(* IEC 61131-3 sources: ctrlx-ai-coding/skills/ctrlx-opcon-engineering/assets/library-examples/inntai/plc/FB_InntaiWireFixture, 4 files *)

(* ---- Close.st ---- *)
METHOD PUBLIC Close : DINT
(* BODY *)
IF ( NOT _opened )
THEN
  AlreadyClosedCalls := AlreadyClosedCalls + 1;
  Close              := -601;
ELSE
  _opened := FALSE;
  Close   := OK;
END_IF

(* ---- Read.st ---- *)
METHOD PUBLIC Read : DINT
VAR_INPUT
  pData        : POINTER TO BYTE;
  DataLen      : SIZE_T;
  rBytesRead   : REFERENCE TO SIZE_T;
  rReadTimeout : REFERENCE TO BOOL;
END_VAR
VAR
  _chunk : UINT;
  _i     : UINT;
END_VAR
(* BODY *)
_chunk := MIN(TO_UINT(DataLen), MIN(_count, 17));
IF ( _chunk > 0 )
THEN
  FOR _i := 0 TO _chunk - 1
  DO
    pData[_i] := _queue[_i];
  END_FOR
  _count := _count - _chunk;
  IF ( _count > 0 )
  THEN
    FOR _i := 0 TO _count - 1
    DO
      _queue[_i] := _queue[_i + _chunk];
    END_FOR
  END_IF
  ReadChunks   := ReadChunks + 1;
  MaxReadChunk := MAX(MaxReadChunk, _chunk);
END_IF
rBytesRead   := _chunk;
rReadTimeout := ( _chunk = 0 );
Read         := OK;

(* ---- Write.st ---- *)
METHOD PUBLIC Write : DINT
VAR_INPUT
  pData         : POINTER TO BYTE;
  DataLen       : SIZE_T;
  rBytesWritten : REFERENCE TO SIZE_T;
END_VAR
VAR
  _bcc : BYTE;
  _i   : UINT;
END_VAR
(* BODY *)
_bcc := 0;
FOR _i := 0 TO TO_UINT(DataLen) - 2
DO
  _bcc := _bcc XOR pData[_i];
END_FOR
WireValid := WireValid AND ( pData[0] = 2 ) AND
             ( pData[DataLen-2] = 3 ) AND ( _bcc = pData[DataLen-1] );
IF ( NOT WireValid )
THEN
  Write := -10009;
  RETURN;
END_IF
IF ( pData[1] = 82 ) AND
   ( pData[2] = 80 )
THEN
  FOR _i := 0 TO SIZEOF(ReplyParameters) - 1
  DO
    _queue[_i] := ReplyParameters[_i];
  END_FOR
  _count := SIZEOF(ReplyParameters);
ELSIF ( pData[1] = 67 ) AND
      ( pData[2] = 83 )
THEN
  CsCalls := CsCalls + 1;
  FOR _i := 0 TO SIZEOF(ReplyBaseline) - 1
  DO
    IF ( FreshOnRead ) THEN
      _queue[_i] := ReplyFresh[_i];
    ELSE
      _queue[_i] := ReplyBaseline[_i];
    END_IF
  END_FOR
  _count := SIZEOF(ReplyBaseline);
ELSE
  FOR _i := 0 TO SIZEOF(ReplyOk) - 1
  DO
    _queue[_i] := ReplyOk[_i];
  END_FOR
  _count   := SIZEOF(ReplyOk);
  _pending := AutoResult AND ( pData[1] = 83 ) AND ( pData[2] = 84 );
  IF ( pData[1] = 83 ) AND ( pData[2] = 84 ) THEN
    StartCalls := StartCalls + 1;
  END_IF
END_IF
IF ( SuppressReply )
THEN
  _count := 0;
END_IF
rBytesWritten := DataLen;
Write         := OK;

(* ---- Open.st ---- *)
METHOD PUBLIC Open : DINT
VAR_INPUT
  BaudRate  : OC_OpconBaseCommonDef.OpconSerialBaudRate;
  DataFrame : OC_OpconBaseCommonDef.OpconSerialDataFrame;
  Handshake : OC_OpconBaseCommonDef.OpconSerialHandshakeType;
END_VAR
(* BODY *)
ConfigurationCorrect :=
(BaudRate = OC_OpconBaseCommonDef.OpconSerialBaudRate.BAUD_9600) AND
(DataFrame = OC_OpconBaseCommonDef.OpconSerialDataFrame.FRAME_8N1) AND
(Handshake = OC_OpconBaseCommonDef.OpconSerialHandshakeType.NO_HANDSHAKE);
IF ( ConfigurationCorrect )
THEN
  IF ( InjectOpenFault )
  THEN
    Open := -21;
  ELSE
    _opened := TRUE;
    Open    := OK;
  END_IF
ELSE
  Open := -1;
END_IF
